(* IEC 61131-3 sources: volt/packages/volt-lsp-iec/test-corpus/twincat-project14/TwinCAT Project14/PLC/Untitled2/Untitled2 Project/GVLs, 1 file *)

(* ---- GVL_PackML.gvl ---- *)
{attribute 'qualified_only'}
VAR_GLOBAL CONSTANT
    UNIT_STATE_TIMEOUT_DEFAULT : TIME := T#10S;
END_VAR
VAR_GLOBAL
END_VAR
